FUNCTION_BLOCK FB_PendantControl
VAR_INPUT
	ipTelescope	: I_RaDecTelescope;
	ipFocus		: I_Focus;
END_VAR
VAR_OUTPUT
END_VAR
VAR
	fbComm			: I_Comm;
	tonComm 		: TON := (PT:=T#5S);
	(*  State Definitions *)
	ipState			: I_PendantState := fbPendantPreInitState;
	ipStateOld		: I_PendantState := fbPendantPreInitState;
	
	fbPendantPreInitState	: FB_PendantPreInitState(THIS);
	fbPendantIdleState 		: FB_PendantIdleState(THIS);
	fbPendantInitState 		: FB_PendantInitState(THIS);
	fbPendantSetHAState		: FB_PendantSetHAState(THIS);
	fbPendantSetDECState	: FB_PendantSetDECState(THIS);
	fbPendantSetFocusState	: FB_PendantSetFocusState(THIS);
	fbPendantErrorState		: FB_PendantErrorState(THIS);
	
	bReady			: BOOL;
	bError			: BOOL;
	bReset			: BOOL;
	nErrorID		: UINT;
	
	(* Set Logic:
		bFastMove:	TRUE (move big step)
					FALSE (move small step)
		bMovePositive:	TRUE +
						FALSE -*)
	bFastMove		: BOOL;
	bMovePositive	: BOOL;
	
	rtrigReset		: R_TRIG;
	rtrigError		: R_TRIG;
	
	(*SEND*)
	fbSendString	: SendString;
	fbSendHex		: SendData;
	eSendErrorID	: ComError_t;
	
	
	(* RECEIVE*)
	fbReceive		: ReceiveString;
	rtrigReceive	: R_TRIG;
	sReceivedString	: STRING;
	sLastReceivedString: STRING;
	bStringReceived	: BOOL;
	bReceiveBusy	: BOOL;
	bReceiveError	: BOOL;
	eReceiveErrorID	: ComError_t;
	bReceiveTimeout	: BOOL;
END_VAR

//	Receive string data:	
fbReceive(
	Prefix:='',
	Suffix:= '',
	Timeout:= T#1MS,
	ReceivedString:= sReceivedString,
	RXbuffer:= RxBufferPendant,
	StringReceived=> bStringReceived,
	Busy=> bReceiveBusy,
	Error=> ,
	RxTimeout=> bReceiveTimeout );

(*Send / Receive Errors? *)
IF fbReceive.Error <> COMERROR_NOERROR THEN
	bError:=TRUE;
	nErrorID		:= fbReceive.Error;
	eReceiveErrorID := fbReceive.Error;
END_IF
IF fbSendString.Error <> COMERROR_NOERROR THEN
	bError:=TRUE;
	nErrorID	:= fbSendString.Error;
	eSendErrorID := fbSendString.Error;
ELSIF fbSendHex.Error <> COMERROR_NOERROR THEN
	bError:=TRUE;
	nErrorID := fbSendHex.Error;
	eSendErrorID := fbSendHex.Error;
END_IF

(* Triggers*)
rtrigReceive(CLK:=bStringReceived);
rtrigReset(CLK:=bReset);
rtrigError(CLK:=bError);

IF rtrigError.Q THEN
	bFastMove := FALSE;
	ipState.FoundError();
ELSIF rtrigReset.Q THEN
	ipState.ResetCommand();
	bReset:=FALSE;
ELSIF rtrigReceive.Q AND NOT bError THEN
	(* INIT *)
	IF sReceivedString = '#' THEN
		ipState.InitCommand();
		
	(* HA *)
	ELSIF sReceivedString = 'û' AND bReady THEN
		(* -, slow*)
		bFastMove := FALSE;
		bMovePositive := FALSE;
		ipState.HaCommand();
	ELSIF sReceivedString = '{' AND bReady THEN
		(* -, fast*)
		bFastMove := TRUE;
		bMovePositive := FALSE;
		ipState.HaCommand();
	ELSIF sReceivedString = 'ý' AND bReady THEN
		(* +, slow*)
		bFastMove := FALSE;
		bMovePositive := TRUE;
		ipState.HaCommand();
	ELSIF sReceivedString = '}' AND bReady THEN
		(* +, fast*)
		bFastMove := TRUE;
		bMovePositive := TRUE;
		ipState.HaCommand();
	
	(* DEC *)
	ELSIF sReceivedString = 'ï' AND bReady THEN
		(* -, slow*)
		bFastMove := FALSE;
		bMovePositive := FALSE;
		ipState.DecCommand();
	ELSIF sReceivedString = 'o' AND bReady THEN
		(* -, fast*)
		bFastMove := TRUE;
		bMovePositive := FALSE;
		ipState.DecCommand();
	ELSIF sReceivedString = '÷' AND bReady THEN
		(* +, slow*)
		bFastMove := FALSE;
		bMovePositive := TRUE;
		ipState.DecCommand();
	ELSIF sReceivedString = 'w' AND bReady THEN
		(* +, fast*)
		bFastMove := TRUE;
		bMovePositive := TRUE;
		ipState.DecCommand();
	
	(* Focus *)
	ELSIF sReceivedString = '¿' AND bReady THEN
		(* -, slow*)
		bFastMove := FALSE;
		bMovePositive := FALSE;
		ipState.FocusCommand();
	ELSIF sReceivedString = '?' AND bReady THEN
		(* -, fast*)
		bFastMove := TRUE;
		bMovePositive := FALSE;
		ipState.FocusCommand();
	ELSIF sReceivedString = 'ß' AND bReady THEN
		(* +, slow*)
		bFastMove := FALSE;
		bMovePositive := TRUE;
		ipState.FocusCommand();
	ELSIF sReceivedString = '_' AND bReady THEN
		(* +, fast*)
		bFastMove := TRUE;
		bMovePositive := TRUE;
		ipState.FocusCommand();
	ELSE
		bFastMove := FALSE;
		ipState.ToIdle();
	END_IF
	
END_IF

ipState.RunState();

PROPERTY _Error : BOOL
GET
_Error := bError;
END_GET
SET
bError:=_Error;
END_SET
END_PROPERTY

PROPERTY _FastMove : BOOL
GET
_FastMove := THIS^.bFastMove;
END_GET
END_PROPERTY

PROPERTY _MovePositive : BOOL
GET
_MovePositive := THIS^.bMovePositive;
END_GET
END_PROPERTY

PROPERTY _Ready : BOOL
GET
_Ready := bReady;
END_GET
SET
bReady := _Ready;
END_SET
END_PROPERTY

PROPERTY Error : BOOL
GET
Error := bError;
END_GET
END_PROPERTY

PROPERTY ErrorID : UINT
GET
ErrorID := nErrorID;
END_GET
END_PROPERTY

//FB_Init is always available implicitly and it is used primarily for initialization.
//The return value is not evaluated. For a specific influence, you can also declare the
//methods explicitly and provide additional code there with the standard initialization
//code. You can evaluate the return value.
METHOD FB_Init: BOOL
VAR_INPUT
    bInitRetains	: BOOL; // TRUE: the retain variables are initialized (reset warm / reset cold)
    bInCopyCode		: BOOL;  // TRUE: the instance will be copied to the copy code afterward (online change)
	comm			: I_Comm;
END_VAR
THIS^.fbComm 				:= comm;
END_METHOD

PROPERTY Reset : BOOL
SET
bReset := Reset;
END_SET
END_PROPERTY

METHOD SetState : BOOL
VAR_INPUT
	newState :I_PendantState;
END_VAR
THIS^.ipState := newState;
END_METHOD

END_FUNCTION_BLOCK

(* stored: Version 1.1.0.1, ProductVersion 3.1.4024.15
   POU FB_PendantControl: Id {31943a3c-0e0b-4aa2-80e9-dadb4d86be37}, SpecialFunc None
   Folder internal properties: Id {a18665bc-e169-47b9-b965-9f2788e06ac9}
   Folder properties: Id {6850b61c-eda9-481c-9524-cd9390cb72ba}
   Property _Error: Id {6593edff-d0b5-41b7-8bc7-58065f448086}
   Get Get: Id {bc020154-760d-4825-8f14-c128881c7e22}
   Set Set: Id {b51dbe17-9c90-44df-adea-ccf9759c05f0}
   Property _FastMove: Id {72cafdb3-ddbc-4b3b-a697-7c53ab685688}
   Get Get: Id {87f3b4e0-9c85-49db-8e48-ba78643e2e06}
   Property _MovePositive: Id {ae64d179-d51b-49a0-810e-4bdae9921153}
   Get Get: Id {8ee045b6-d5ee-4db5-b9dc-cb8d6dc97da2}
   Property _Ready: Id {6219a3da-e3d8-44a9-b851-742f91d2d543}
   Get Get: Id {35c150dd-44cc-45f8-b83d-10d48a514af0}
   Set Set: Id {ac77bf06-0f7e-48a8-a327-c7d65024c7ea}
   Property Error: Id {8bfc8674-e993-417b-9a6d-81cdaeebc0e0}
   Get Get: Id {40fb6eb4-7078-4cd9-9b43-da41422a828f}
   Property ErrorID: Id {2176f647-c267-4999-83ee-92a6d6d1ebd3}
   Get Get: Id {3fecda0a-f327-4f18-9714-138ac84670e7}
   Method FB_Init: Id {7299abf0-bea5-41f3-9d4e-3091c390ab64}
   Property Reset: Id {45d22cd5-17ee-46bf-9f0b-8a5cb1bbc7ed}
   Set Set: Id {3432f7db-0aa8-4e51-b308-169338550f01}
   Method SetState: Id {a8389db5-f741-4ceb-b61b-f12dece5de1d} *)
